(* IEC 61131-3 sources: tsplc/examples/bottling-line/raw-st/src/common, 1 file *)

(* ---- F_Clamp.st ---- *)
FUNCTION F_Clamp : INT
VAR_INPUT
	Value : INT;
	Low : INT;
	High : INT;
END_VAR
F_Clamp := MIN(MAX(Value, Low), High);
END_FUNCTION
